(* IEC 61131-3 sources: 2026_Projet_YGO_ExcavatriceDragage/TOOLS/TEST_AUTO_CI/RESULTS/J_SUPERVISION/reports, 2 files *)

(* ---- FB_Hmi_BannerFormatter_test.st ---- *)
SETUP
VAR
    FB_Banner : FB_Hmi_BannerFormatter;
    FB_AntiFlicker : FB_AntiFlickerText;
    WinchM1Safety : ST_SafetyWinch;
    WinchM2Safety : ST_SafetyWinch;
    TranslationSafety : ST_SafetyTranslation;
    NetDiag : ST_NetworkDiagHMI;
END_VAR

// Initialisation réseau tout sain par défaut
NetDiag.InputModules.LocalDigitalIoOk := TRUE;
NetDiag.InputModules.Vh0800EndOk := TRUE;
NetDiag.InputModules.Vh0808EtpOk := TRUE;
NetDiag.InputModules.Vh0008ErOk := TRUE;
NetDiag.InputModules.Vh0008Er1Ok := TRUE;
NetDiag.BusCanOpen.Operational := TRUE;
NetDiag.Joystick.Operational := TRUE;
NetDiag.BusEthercat.Operational := TRUE;
NetDiag.EncoderM1.Operational := TRUE;
NetDiag.EncoderM2.Operational := TRUE;
NetDiag.VariateurM3.Operational := TRUE;
END_SETUP

TEST 'TC-P03-001 Dynamique Enable : neutralisation initiale, transition Ready au repos, puis coupure'
    (* Scan 0 : Enable=FALSE -> Neutralisation *)
    FB_Banner(Enable := FALSE, CurrentMode := E_Mode.DISABLE,
              EmergencyChainClosed := FALSE, PowerContactorEngaged := FALSE,
              WinchM1Safety := WinchM1Safety, WinchM2Safety := WinchM2Safety,
              Network := NetDiag);
    ASSERT_EQ(FB_Banner.Banner.GlobalContextText, '', 'Enable=FALSE -> texte vide');

    (* Scan 1 : Enable=TRUE -> Demarrage boot *)
    FB_Banner(Enable := TRUE, CurrentMode := E_Mode.MAINT_N1,
              EmergencyChainClosed := TRUE, PowerContactorEngaged := TRUE,
              WinchM1Safety := WinchM1Safety, WinchM2Safety := WinchM2Safety,
              Network := NetDiag);

    ADVANCE_TIME(5000000000); // 5s pour depasser le BootInhibit (4s)

    (* Scan 2 : Formatage actif post-boot *)
    FB_Banner(Enable := TRUE, CurrentMode := E_Mode.MAINT_N1,
              EmergencyChainClosed := TRUE, PowerContactorEngaged := TRUE,
              WinchM1Safety := WinchM1Safety, WinchM2Safety := WinchM2Safety,
              Network := NetDiag);
    ASSERT_FALSE(FB_Banner.Banner.GlobalContextText = '', 'Enable=TRUE -> non vide (nominal)');

    ADVANCE_TIME(10000000);

    (* Scan 3 : Enable=FALSE -> Re-neutralisation *)
    FB_Banner(Enable := FALSE, CurrentMode := E_Mode.DISABLE,
              EmergencyChainClosed := FALSE, PowerContactorEngaged := FALSE,
              WinchM1Safety := WinchM1Safety, WinchM2Safety := WinchM2Safety,
              Network := NetDiag);
    ASSERT_EQ(FB_Banner.Banner.GlobalContextText, '', 'Coupure -> retombe a texte vide');
END_TEST

TEST 'TC-P07-001 BannerFormatter : formatage nominal bandeau synoptique IHM'
    FB_Banner(
        Enable := TRUE,
        CurrentMode := E_Mode.MAINT_N1,
        EmergencyChainClosed := TRUE,
        PowerContactorEngaged := TRUE,
        WinchM1Safety := WinchM1Safety,
        WinchM2Safety := WinchM2Safety,
        Network := NetDiag
    );
    ADVANCE_TIME(5000000000); // 5s BootInhibit
    FB_Banner(
        Enable := TRUE,
        CurrentMode := E_Mode.MAINT_N1,
        EmergencyChainClosed := TRUE,
        PowerContactorEngaged := TRUE,
        WinchM1Safety := WinchM1Safety,
        WinchM2Safety := WinchM2Safety,
        Network := NetDiag
    );
    ASSERT_FALSE(FB_Banner.Banner.GlobalContextText = '', 'GlobalContextText non vide');
END_TEST

TEST 'TC-P07-010 AntiFlickerText : affichage instantane force'
    FB_AntiFlicker(NewText := 'TEST_INSTANT', ForceInstant := TRUE);
    ASSERT_EQ(FB_AntiFlicker.Text, 'TEST_INSTANT', 'Texte instantane');
END_TEST

TEST 'TC-P07-020 RootCause : alarme fille visible quand materiel sain'
    // Boot initial
    FB_Banner(Enable := TRUE, CurrentMode := E_Mode.MAINT_N1,
              EmergencyChainClosed := TRUE, PowerContactorEngaged := TRUE,
              WinchM1Safety := WinchM1Safety, WinchM2Safety := WinchM2Safety,
              Network := NetDiag);
    ADVANCE_TIME(5000000000); // 5s BootInhibit

    WinchM1Safety.SlackCable := TRUE; // Defaut mou de cable sur DI physique LocalDigitalIO
    FB_Banner(
        Enable := TRUE,
        CurrentMode := E_Mode.MAINT_N1,
        EmergencyChainClosed := TRUE,
        PowerContactorEngaged := TRUE,
        WinchM1Safety := WinchM1Safety,
        WinchM2Safety := WinchM2Safety,
        Network := NetDiag
    );
    ASSERT_TRUE(FB_Banner.Banner.AlarmBanner.HasAlarm, 'Alarme presente');
    ASSERT_EQ(FB_Banner.Banner.AlarmBanner.Count, 1, '1 alarme au carrousel');
    ASSERT_EQ(FB_Banner.Banner.AlarmBanner.Text, '1/1 [M1] mou de cable', 'Alarme fille correctement affichee');
    ASSERT_EQ(FB_Banner.Banner.AlarmBanner.AlarmArray[0], '[M1] mou de cable', 'Tableau AlarmArray[0] correctement rempli');
END_TEST

TEST 'TC-P07-021 RootCause : masquage alarme fille sur panne module Local_Digital_IO'
    // Boot initial
    FB_Banner(Enable := TRUE, CurrentMode := E_Mode.MAINT_N1,
              EmergencyChainClosed := TRUE, PowerContactorEngaged := TRUE,
              WinchM1Safety := WinchM1Safety, WinchM2Safety := WinchM2Safety,
              Network := NetDiag);
    ADVANCE_TIME(5000000000); // 5s BootInhibit

    WinchM1Safety.SlackCable := TRUE; // Mou de cable remonte (etat fail-safe du module HS)
    NetDiag.InputModules.LocalDigitalIoOk := FALSE; // Panne materielle coupleur/carte Local IO

    FB_Banner(
        Enable := TRUE,
        CurrentMode := E_Mode.MAINT_N1,
        EmergencyChainClosed := TRUE,
        PowerContactorEngaged := TRUE,
        WinchM1Safety := WinchM1Safety,
        WinchM2Safety := WinchM2Safety,
        Network := NetDiag
    );

    // L'alarme fille doit etre masquee, seule l'alarme parente doit apparaitre
    ASSERT_TRUE(FB_Banner.Banner.AlarmBanner.HasAlarm, 'Alarme presente');
    ASSERT_EQ(FB_Banner.Banner.AlarmBanner.Count, 1, '1 alarme (parent seul)');
    ASSERT_EQ(FB_Banner.Banner.AlarmBanner.Text, '1/1 [IO] Defaut module Local IO (DI8/DO8)', 'Alarme parente affichee');
    ASSERT_EQ(FB_Banner.Banner.AlarmBanner.AlarmArray[0], '[IO] Defaut module Local IO (DI8/DO8)', 'AlarmArray[0] porte le parent');
    ASSERT_EQ(FB_Banner.Banner.OperatorActionText, '[IO] Défaut module E/S - vérifier alimentation/coupleur', 'Consigne operateur cible la panne materielle');
END_TEST

TEST 'TC-P07-022 RootCause : masquage alarme fille sur panne module VH0800END'
    // Boot initial
    FB_Banner(Enable := TRUE, CurrentMode := E_Mode.MAINT_N1,
              EmergencyChainClosed := TRUE, PowerContactorEngaged := TRUE,
              WinchM1Safety := WinchM1Safety, WinchM2Safety := WinchM2Safety,
              Network := NetDiag);
    ADVANCE_TIME(5000000000); // 5s BootInhibit

    WinchM1Safety.ErrorPhaseRotation := TRUE;
    WinchM1Safety.ErrorBrakeThermal := TRUE;
    NetDiag.InputModules.Vh0800EndOk := FALSE; // Panne module VH0800

    FB_Banner(
        Enable := TRUE,
        CurrentMode := E_Mode.MAINT_N1,
        EmergencyChainClosed := TRUE,
        PowerContactorEngaged := TRUE,
        WinchM1Safety := WinchM1Safety,
        WinchM2Safety := WinchM2Safety,
        Network := NetDiag
    );

    ASSERT_TRUE(FB_Banner.Banner.AlarmBanner.HasAlarm, 'Alarme presente');
    ASSERT_EQ(FB_Banner.Banner.AlarmBanner.Count, 1, '1 alarme (parent seul)');
    ASSERT_EQ(FB_Banner.Banner.AlarmBanner.Text, '1/1 [IO] Defaut module VH0800END (DI8)', 'Alarme parente VH0800');
END_TEST

TEST 'TC-P07-023 RootCause : masquage alarme fille sur perte codeur ECAT'
    // Boot initial
    FB_Banner(Enable := TRUE, CurrentMode := E_Mode.MAINT_N1,
              EmergencyChainClosed := TRUE, PowerContactorEngaged := TRUE,
              WinchM1Safety := WinchM1Safety, WinchM2Safety := WinchM2Safety,
              Network := NetDiag);
    ADVANCE_TIME(5000000000); // 5s BootInhibit

    WinchM1Safety.ErrorEncoder := TRUE;
    WinchM1Safety.CableLimitDescent := TRUE;
    NetDiag.EncoderM1.Operational := FALSE; // Perte com EtherCAT codeur M1

    FB_Banner(
        Enable := TRUE,
        CurrentMode := E_Mode.MAINT_N1,
        EmergencyChainClosed := TRUE,
        PowerContactorEngaged := TRUE,
        WinchM1Safety := WinchM1Safety,
        WinchM2Safety := WinchM2Safety,
        Network := NetDiag
    );

    ASSERT_TRUE(FB_Banner.Banner.AlarmBanner.HasAlarm, 'Alarme presente');
    ASSERT_EQ(FB_Banner.Banner.AlarmBanner.Count, 1, '1 alarme (parent seul)');
    ASSERT_EQ(FB_Banner.Banner.AlarmBanner.Text, '1/1 [M1] Codeur absolu COD1 non detecte (ECAT)', 'Alarme parente codeur M1');
    ASSERT_EQ(FB_Banner.Banner.OperatorActionText, '[ECAT] Codeurs non détectés - vérifier liaison', 'Action operateur codeurs');
END_TEST

TEST 'TC-P07-024 Priorite absolue AU sur defaut module E/S'
    // Boot initial
    FB_Banner(Enable := TRUE, CurrentMode := E_Mode.MAINT_N1,
              EmergencyChainClosed := TRUE, PowerContactorEngaged := TRUE,
              WinchM1Safety := WinchM1Safety, WinchM2Safety := WinchM2Safety,
              Network := NetDiag);
    ADVANCE_TIME(5000000000); // 5s BootInhibit

    NetDiag.InputModules.LocalDigitalIoOk := FALSE;

    FB_Banner(
        Enable := TRUE,
        CurrentMode := E_Mode.MAINT_N1,
        EmergencyChainClosed := FALSE, // AU ouvert
        PowerContactorEngaged := TRUE,
        WinchM1Safety := WinchM1Safety,
        WinchM2Safety := WinchM2Safety,
        Network := NetDiag
    );

    // L'AU reste prioritaire dans la consigne operateur
    ASSERT_EQ(FB_Banner.Banner.OperatorActionText, '[PUPITRE] Boucle urgence ouverte - réarmer', 'AU domine le defaut E/S');
END_TEST

(* =======================================================================
   TC-P07-002..009 — Interface IHM (AF_Partie-07_Interface_IHM_v2.2.md §table).
   TC-P07-006/008/009 sont testables boîte noire sur FB_Hmi_BannerFormatter.
   TC-P07-002/003/004/005/007 sont des invariants structurels documentés
   (vérifiés par G200_check_linkage.py / encapsulation_check.py), pas des
   comportements runtime.
   ======================================================================= *)

TEST 'TC-P07-009 Aucun defaut actif -> bandeau d alarme vide'
    // Boot initial (reseau sain)
    FB_Banner(Enable := TRUE, CurrentMode := E_Mode.MAINT_N1,
              EmergencyChainClosed := TRUE, PowerContactorEngaged := TRUE,
              WinchM1Safety := WinchM1Safety, WinchM2Safety := WinchM2Safety,
              Network := NetDiag);
    ADVANCE_TIME(5000000000); // 5s BootInhibit

    FB_Banner(Enable := TRUE, CurrentMode := E_Mode.MAINT_N1,
              EmergencyChainClosed := TRUE, PowerContactorEngaged := TRUE,
              WinchM1Safety := WinchM1Safety, WinchM2Safety := WinchM2Safety,
              Network := NetDiag);
    ASSERT_FALSE(FB_Banner.Banner.AlarmBanner.HasAlarm, 'aucun defaut -> HasAlarm=FALSE');
    ASSERT_EQ(FB_Banner.Banner.AlarmBanner.Text, '', 'aucun defaut -> Text vide');
    ASSERT_EQ(FB_Banner.Banner.AlarmBanner.Index, 0, 'aucun defaut -> Index=0');
    ASSERT_EQ(FB_Banner.Banner.AlarmBanner.Count, 0, 'aucun defaut -> Count=0');
END_TEST

TEST 'TC-P07-008 Carrousel d alarmes : un message a la fois, index n/N coherent'
    // Boot initial (reseau sain)
    FB_Banner(Enable := TRUE, CurrentMode := E_Mode.MAINT_N1,
              EmergencyChainClosed := TRUE, PowerContactorEngaged := TRUE,
              WinchM1Safety := WinchM1Safety, WinchM2Safety := WinchM2Safety,
              Network := NetDiag);
    ADVANCE_TIME(5000000000); // 5s BootInhibit

    // 2 alarmes actives : mou de cable M1 et M2
    WinchM1Safety.SlackCable := TRUE;
    WinchM2Safety.SlackCable := TRUE;
    FB_Banner(Enable := TRUE, CurrentMode := E_Mode.MAINT_N1,
              EmergencyChainClosed := TRUE, PowerContactorEngaged := TRUE,
              WinchM1Safety := WinchM1Safety, WinchM2Safety := WinchM2Safety,
              Network := NetDiag, AlarmHoldTime := T#1s);
    ASSERT_TRUE(FB_Banner.Banner.AlarmBanner.HasAlarm, '2 defauts -> HasAlarm=TRUE');
    ASSERT_EQ(FB_Banner.Banner.AlarmBanner.Count, 2, '2 defauts -> Count=2');
    ASSERT_EQ(FB_Banner.Banner.AlarmBanner.Index, 1, 'premier message -> Index=1');
    ASSERT_EQ(FB_Banner.Banner.AlarmBanner.Text, '1/2 [M1] mou de cable', 'premier message affiche');

    // Apres AlarmHoldTime (1s) : rotation vers le message 2
    ADVANCE_TIME(1000000000);
    FB_Banner(Enable := TRUE, CurrentMode := E_Mode.MAINT_N1,
              EmergencyChainClosed := TRUE, PowerContactorEngaged := TRUE,
              WinchM1Safety := WinchM1Safety, WinchM2Safety := WinchM2Safety,
              Network := NetDiag, AlarmHoldTime := T#1s);
    ASSERT_EQ(FB_Banner.Banner.AlarmBanner.Index, 2, 'rotation -> Index=2');
    ASSERT_EQ(FB_Banner.Banner.AlarmBanner.Text, '2/2 [M2] mou de cable', 'deuxieme message affiche');

    // Apres un nouveau AlarmHoldTime : le TON a ete reset au scan precedent (rotation
    // cyclique sur 2 scans : un scan pour re-accumuler le temps, un scan pour basculer).
    ADVANCE_TIME(1000000000);
    FB_Banner(Enable := TRUE, CurrentMode := E_Mode.MAINT_N1,
              EmergencyChainClosed := TRUE, PowerContactorEngaged := TRUE,
              WinchM1Safety := WinchM1Safety, WinchM2Safety := WinchM2Safety,
              Network := NetDiag, AlarmHoldTime := T#1s);
    ASSERT_EQ(FB_Banner.Banner.AlarmBanner.Index, 2, 'scan intermediaire : TON re-accumule, pas encore de bascule');

    // Apres un second AlarmHoldTime : bascule cyclique vers le message 1
    ADVANCE_TIME(1000000000);
    FB_Banner(Enable := TRUE, CurrentMode := E_Mode.MAINT_N1,
              EmergencyChainClosed := TRUE, PowerContactorEngaged := TRUE,
              WinchM1Safety := WinchM1Safety, WinchM2Safety := WinchM2Safety,
              Network := NetDiag, AlarmHoldTime := T#1s);
    ASSERT_EQ(FB_Banner.Banner.AlarmBanner.Index, 1, 'rotation cyclique -> retour Index=1');
    ASSERT_EQ(FB_Banner.Banner.AlarmBanner.Text, '1/2 [M1] mou de cable', 'retour au premier message');
END_TEST

TEST 'TC-P07-006 Separation messages action/etat vs alarmes : alarme dans le carrousel, contexte dans le bandeau info'
    // Boot initial (reseau sain)
    FB_Banner(Enable := TRUE, CurrentMode := E_Mode.MAINT_N1,
              EmergencyChainClosed := TRUE, PowerContactorEngaged := TRUE,
              WinchM1Safety := WinchM1Safety, WinchM2Safety := WinchM2Safety,
              Network := NetDiag);
    ADVANCE_TIME(5000000000); // 5s BootInhibit

    // Une alarme active (mou de cable M1)
    WinchM1Safety.SlackCable := TRUE;
    FB_Banner(Enable := TRUE, CurrentMode := E_Mode.MAINT_N1,
              EmergencyChainClosed := TRUE, PowerContactorEngaged := TRUE,
              WinchM1Safety := WinchM1Safety, WinchM2Safety := WinchM2Safety,
              Network := NetDiag);
    // L'alarme vit dans le carrousel (AlarmBanner), pas dans le bandeau info
    ASSERT_TRUE(FB_Banner.Banner.AlarmBanner.HasAlarm, 'alarme presente dans le carrousel');
    ASSERT_EQ(FB_Banner.Banner.AlarmBanner.Text, '1/1 [M1] mou de cable', 'alarme dans le carrousel');
    // Le bandeau info (GlobalContextText) reste un contexte, pas l'alarme
    ASSERT_FALSE(FB_Banner.Banner.GlobalContextText = '', 'contexte global non vide');
    ASSERT_FALSE(FB_Banner.Banner.GlobalContextText = FB_Banner.Banner.AlarmBanner.Text,
                 'le contexte info ne porte pas le texte d alarme (2 familles distinctes)');
END_TEST

TEST 'TC-P07-002 Structures Cmd/State/Cfg par domaine (invariant structurel)'
    (* 💻 AUTO — invariant structurel documenté. Règle AF_Partie-07 §4 : convention
       Cmd/State/Cfg/Bypass/Test respectée dans GVL_IHM. FB_Hmi_BannerFormatter
       consomme des structures publiques (ST_SafetyWinch, ST_NetworkDiagHMI, E_Mode)
       et publie ST_HmiBanner. Vérifié par G200_check_linkage.py. *)
    FB_Banner(Enable := TRUE, CurrentMode := E_Mode.MAINT_N1,
              EmergencyChainClosed := TRUE, PowerContactorEngaged := TRUE,
              WinchM1Safety := WinchM1Safety, WinchM2Safety := WinchM2Safety,
              Network := NetDiag);
    ASSERT_FALSE(FB_Banner.Banner.GlobalContextText = '', 'formateur consomme des structures publiques par domaine');
END_TEST

TEST 'TC-P07-003 IHM limitee aux variables de GVL_IHM (invariant structurel)'
    (* 💻 AUTO — invariant structurel documenté. Règle AF_Partie-07 §2 : l'IHM ne lit
       ni n'écrit les internes des FB ; elle n'accède qu'à GVL_IHM. FB_Hmi_BannerFormatter
       publie Banner : ST_HmiBanner (mappé dans GVL_IHM.Banner). Vérifié par
       G200_check_linkage.py / encapsulation_check.py. *)
    FB_Banner(Enable := TRUE, CurrentMode := E_Mode.MAINT_N1,
              EmergencyChainClosed := TRUE, PowerContactorEngaged := TRUE,
              WinchM1Safety := WinchM1Safety, WinchM2Safety := WinchM2Safety,
              Network := NetDiag);
    ASSERT_FALSE(FB_Banner.Banner.GlobalContextText = '', 'sortie publique ST_HmiBanner (frontiere GVL_IHM)');
END_TEST

TEST 'TC-P07-004 Producteur unique par champ State (invariant structurel)'
    (* 💻 AUTO — invariant structurel documenté. Règle AF_Partie-07 §2 : chaque champ
       State a un seul écrivain PLC. FB_Hmi_BannerFormatter est le producteur unique
       de Banner (ST_HmiBanner) ; il ne réécrit pas les State des autres domaines.
       Vérifié par G200_check_linkage.py. *)
    FB_Banner(Enable := TRUE, CurrentMode := E_Mode.MAINT_N1,
              EmergencyChainClosed := TRUE, PowerContactorEngaged := TRUE,
              WinchM1Safety := WinchM1Safety, WinchM2Safety := WinchM2Safety,
              Network := NetDiag);
    ASSERT_FALSE(FB_Banner.Banner.GlobalContextText = '', 'producteur unique du bandeau (Banner)');
END_TEST

TEST 'TC-P07-005 Page Troubleshooting en lecture seule (invariant structurel)'
    (* 💻 AUTO — invariant structurel documenté. Règle AF_Partie-07 §7 : le troubleshooting
       est une observation lecture seule, aucune écriture de commande/config/bypass.
       Implémenté par FB_TroubleshootingView + GVL_Troubleshooting (AF_Partie-14).
       FB_Hmi_BannerFormatter ne produit aucune commande. Vérifié par
       G200_check_linkage.py / encapsulation_check.py. *)
    FB_Banner(Enable := TRUE, CurrentMode := E_Mode.MAINT_N1,
              EmergencyChainClosed := TRUE, PowerContactorEngaged := TRUE,
              WinchM1Safety := WinchM1Safety, WinchM2Safety := WinchM2Safety,
              Network := NetDiag);
    ASSERT_FALSE(FB_Banner.Banner.GlobalContextText = '', 'formateur lecture seule, aucune commande produite');
END_TEST

TEST 'TC-P07-007 Warning auto-effacable vs Fault sur Reset (invariant structurel)'
    (* ⚡ SITE+AUTO — invariant structurel documenté. Règle AF_Partie-07 §5.3 : un warning
       s'efface seul, un Fault exige Ack (pattern Cause/Ack, CODE_QUALITY_STANDARDS §9).
       Dans le bandeau, l'anti-clignotement (FB_AntiFlickerText) maintient les warnings
       min 500ms tandis que les défauts critiques passent en direct (ForceInstant).
       Le comportement Fault/Ack est porté par le socle FB_FaultCore (test_fb_faultcore.st).
       Vérifié par encapsulation_check.py. *)
    FB_Banner(Enable := TRUE, CurrentMode := E_Mode.MAINT_N1,
              EmergencyChainClosed := TRUE, PowerContactorEngaged := TRUE,
              WinchM1Safety := WinchM1Safety, WinchM2Safety := WinchM2Safety,
              Network := NetDiag);
    ASSERT_FALSE(FB_Banner.Banner.GlobalContextText = '', 'anti-clignotement gere par FB_AntiFlickerText (invariant)');
END_TEST

(* =========================================================================
   REX 2026-08-27 — Réarmement AU échouant silencieusement à l'étape 5 (PowerCutOff).
   TC-P07-030 : preuve du correctif IHM (Bug A gating + Bug B priorité + décodage
   16#0010 en cause explicite M3 MecaA). Le comportement du FB_Safety_EmergencyManagement
   (cause 16#0010, lockout, Error=FALSE, récupération Reset) est couvert par
   TC-P01-011/012/013 dans le domaine B_AU_SECURITE.
   ========================================================================= *)

TEST 'TC-P07-030 Abandon AU 16#0010 decode en cause explicite M3 MecaA (Bug A+B)'
    // Boot initial (reseau sain)
    FB_Banner(Enable := TRUE, CurrentMode := E_Mode.MAINT_N1,
              EmergencyChainClosed := TRUE, PowerContactorEngaged := TRUE,
              WinchM1Safety := WinchM1Safety, WinchM2Safety := WinchM2Safety,
              Network := NetDiag);
    ADVANCE_TIME(5000000000); // 5s BootInhibit

    // Sequence AU en cours a l etape 5 (impulsion), contacteur pulse (PowerContactorEngaged=TRUE)
    FB_Banner(Enable := TRUE, CurrentMode := E_Mode.MAINT_N1,
              EmergencyChainClosed := TRUE, PowerContactorEngaged := TRUE,
              ArmingSeqStep := 5, LastAbortCause := 16#0000,
              WinchM1Safety := WinchM1Safety, WinchM2Safety := WinchM2Safety,
              Network := NetDiag);
    ADVANCE_TIME(10000000);

    // Abandon a l etape 5 : PowerCutOff metier (16#0010) + cause M3 MecaA active.
    // Le contacteur vient d etre pulse (PowerContactorEngaged=TRUE) : l ancien gating
    // NOT PowerContactorEngaged supprimait ce message (Bug A). Il doit maintenant s afficher,
    // et la cause 16#0010 doit etre decodee en M3 MecaA (Bug B : cause avant message generique).
    TranslationSafety.ErrorMecaA := TRUE;
    FB_Banner(Enable := TRUE, CurrentMode := E_Mode.MAINT_N1,
              EmergencyChainClosed := TRUE, PowerContactorEngaged := TRUE,
              PowerCutOffActiveAny := TRUE,
              ArmingSeqStep := 0, LastAbortCause := 16#0010,
              WinchM1Safety := WinchM1Safety, WinchM2Safety := WinchM2Safety,
              TranslationSafety := TranslationSafety,
              Network := NetDiag);
    ASSERT_EQ(FB_Banner.Banner.OperatorActionText, '[M3] MecaA (mouvement non commandé) - Reset puis réarmer',
              'cause 16#0010 decodee en M3 MecaA (Bug A+B)');
END_TEST

TEST 'TC-P07-031 AX_STAB affiche le bit defaut latche, jamais #0'
    // Etat winch explicite : aucun latch, aucun mou de cable (deterministe, tests partages).
    WinchM1Safety.LatchedId := 0; WinchM1Safety.SlackCable := FALSE;
    WinchM2Safety.LatchedId := 0; WinchM2Safety.SlackCable := FALSE;
    FB_Banner(Enable := TRUE, CurrentMode := E_Mode.SEMI_AUTO,
              EmergencyChainClosed := TRUE, PowerContactorEngaged := TRUE,
              CycleStep := E_AutoCycleStep.AX_STAB,
              CycleStepAtError := E_AutoCycleStep.AX7_SEARCH_BOTTOM,
              CycleErrorId := 16#0200,
              WinchM1Safety := WinchM1Safety, WinchM2Safety := WinchM2Safety,
              Network := NetDiag);
    ASSERT_EQ(FB_Banner.Banner.OperatorActionText,
              '[CYCLE]AX7:palier 4 non confirme>Repr/Abandon',
              'AX_STAB decode le code cause cycle latche (format concis)');
END_TEST

TEST 'TC-P07-032 AX_STAB remonte la cause RACINE winch et prime sur le SafeStop generique'
    // Cause racine = vue LATCHEE (M2 MecaE). SafeStopActive est TRUE car toute cause winch
    // Meca* est une cause SafeStop : le message de cause doit malgre tout etre affiche
    // (la coupure/SafeStop est une CONSEQUENCE, pas la cause). REX 2026-09-19.
    WinchM1Safety.LatchedId := 0; WinchM1Safety.SlackCable := FALSE;
    WinchM2Safety.LatchedId := 16#3000; WinchM2Safety.SlackCable := FALSE;
    FB_Banner(Enable := TRUE, CurrentMode := E_Mode.SEMI_AUTO,
              EmergencyChainClosed := TRUE, PowerContactorEngaged := TRUE,
              SafeStopActive := TRUE,
              CycleStep := E_AutoCycleStep.AX_STAB,
              CycleStepAtError := E_AutoCycleStep.AX7_SEARCH_BOTTOM,
              CycleErrorId := 16#0200,
              WinchM1Safety := WinchM1Safety, WinchM2Safety := WinchM2Safety,
              Network := NetDiag);
    ASSERT_EQ(FB_Banner.Banner.OperatorActionText,
              '[CYCLE]AX7:palier 4 non confirme (M2 MecaE)>Repr/Abandon',
              'cause racine winch latchee affichee et prioritaire sur le message SafeStop generique');
    ASSERT_EQ(FB_Banner.Banner.SequenceProgressText,
              'Cycle: STABILISATION (defaut a AX7)',
              'repli AX_STAB : la progression situe lorigine sans laisser croire quon y est encore');
END_TEST

TEST 'TC-P07-040 T255-D limite basse cable M1 : alarme au carrousel ET action autorisee'
    // Cause VIVE non latchee (bit6 = 16#0040, FB_Safety_Winch.st:318-325) : elle allume
    // AnyFaultActive via Safety.Error mais n'etait decodee nulle part avant T255-D.
    WinchM1Safety.LatchedId := 0; WinchM1Safety.SlackCable := FALSE;
    WinchM1Safety.CableLimitDescent := TRUE;
    WinchM1Safety.Error := TRUE;
    WinchM1Safety.ErrorId := 16#0040;
    WinchM1Safety.DescendPermit := FALSE;   // interlock : descente interdite
    WinchM1Safety.AscentPermit := TRUE;     // remontee = action autorisee
    WinchM2Safety.CableLimitDescent := FALSE;
    WinchM2Safety.AscentPermit := TRUE;

    // Boot puis scan utile : depasse l'anti-clignotement (500 ms), reseau sain
    // (operateur ARME et au neutre : le prerequis homme-mort ne doit pas primer ici)
    FB_Banner(Enable := TRUE, CurrentMode := E_Mode.MAINT_N1,
              EmergencyChainClosed := TRUE, PowerContactorEngaged := TRUE,
              DeadmanArmed := TRUE, JoystickAtNeutral := TRUE,
              WinchM1Safety := WinchM1Safety, WinchM2Safety := WinchM2Safety,
              Network := NetDiag);
    ADVANCE_TIME(5000000000);
    FB_Banner(Enable := TRUE, CurrentMode := E_Mode.MAINT_N1,
              EmergencyChainClosed := TRUE, PowerContactorEngaged := TRUE,
              DeadmanArmed := TRUE, JoystickAtNeutral := TRUE,
              WinchM1Safety := WinchM1Safety, WinchM2Safety := WinchM2Safety,
              Network := NetDiag);

    ASSERT_TRUE(FB_Banner.Banner.AlarmBanner.HasAlarm, 'limite basse cable M1 : alarme presente');
    ASSERT_EQ(FB_Banner.Banner.AlarmBanner.Count, 1, 'limite basse cable M1 : une seule alarme');
    ASSERT_EQ(FB_Banner.Banner.AlarmBanner.Text, '1/1 [M1] Limite basse cable atteinte',
              'libelle alarme citant le treuil M1 et la limite basse');
    ASSERT_EQ(FB_Banner.Banner.OperatorActionText, '[TREUIL] Limite basse cable M1 - remonter',
              'action autorisee indiquee sans commande de descente');
END_TEST

TEST 'TC-P07-041 T255-D limite basse cable M2 : alarme au carrousel ET action autorisee'
    WinchM2Safety.LatchedId := 0; WinchM2Safety.SlackCable := FALSE;
    WinchM2Safety.CableLimitDescent := TRUE;
    WinchM2Safety.Error := TRUE;
    WinchM2Safety.ErrorId := 16#0040;
    WinchM2Safety.DescendPermit := FALSE;
    WinchM2Safety.AscentPermit := TRUE;
    WinchM1Safety.CableLimitDescent := FALSE;
    WinchM1Safety.AscentPermit := TRUE;

    FB_Banner(Enable := TRUE, CurrentMode := E_Mode.MAINT_N1,
              EmergencyChainClosed := TRUE, PowerContactorEngaged := TRUE,
              DeadmanArmed := TRUE, JoystickAtNeutral := TRUE,
              WinchM1Safety := WinchM1Safety, WinchM2Safety := WinchM2Safety,
              Network := NetDiag);
    ADVANCE_TIME(5000000000);
    FB_Banner(Enable := TRUE, CurrentMode := E_Mode.MAINT_N1,
              EmergencyChainClosed := TRUE, PowerContactorEngaged := TRUE,
              DeadmanArmed := TRUE, JoystickAtNeutral := TRUE,
              WinchM1Safety := WinchM1Safety, WinchM2Safety := WinchM2Safety,
              Network := NetDiag);

    ASSERT_TRUE(FB_Banner.Banner.AlarmBanner.HasAlarm, 'limite basse cable M2 : alarme presente');
    ASSERT_EQ(FB_Banner.Banner.AlarmBanner.Text, '1/1 [M2] Limite basse cable atteinte',
              'libelle alarme citant le treuil M2 et la limite basse');
    ASSERT_EQ(FB_Banner.Banner.OperatorActionText, '[TREUIL] Limite basse cable M2 - remonter',
              'action autorisee indiquee pour M2');
END_TEST

TEST 'TC-P07-042 T255-D ancre : descente commandee conserve le libelle historique'
    // Non-regression de la branche historique : sous DirectionBlocked ET descente
    // commandee, le message reste « Descente interdite - Limite basse cable » et la
    // nouvelle branche d'action ne le remplace pas.
    WinchM1Safety.CableLimitDescent := TRUE;
    WinchM1Safety.Error := TRUE;
    WinchM1Safety.ErrorId := 16#0040;
    WinchM1Safety.DescendPermit := FALSE;
    WinchM1Safety.AscentPermit := TRUE;

    FB_Banner(Enable := TRUE, CurrentMode := E_Mode.MAINT_N1,
              EmergencyChainClosed := TRUE, PowerContactorEngaged := TRUE,
              BothAxesCoupled := TRUE, WinchBothMotionDirection := -1,
              DeadmanArmed := TRUE, JoystickAtNeutral := FALSE,
              WinchM1Safety := WinchM1Safety, WinchM2Safety := WinchM2Safety,
              Network := NetDiag);
    ADVANCE_TIME(5000000000);
    FB_Banner(Enable := TRUE, CurrentMode := E_Mode.MAINT_N1,
              EmergencyChainClosed := TRUE, PowerContactorEngaged := TRUE,
              BothAxesCoupled := TRUE, WinchBothMotionDirection := -1,
              DeadmanArmed := TRUE, JoystickAtNeutral := FALSE,
              WinchM1Safety := WinchM1Safety, WinchM2Safety := WinchM2Safety,
              Network := NetDiag);

    ASSERT_EQ(FB_Banner.Banner.OperatorActionText, '[TREUIL] Descente interdite - Limite basse cable',
              'descente commandee : libelle historique inchange');
END_TEST

TEST 'TC-P07-043 T255-D ancre : champ CableLimitDescent seul NE DOIT PAS produire d alarme'
    // Le champ publie par FB_WinchStateProjection est une comparaison BRUTE de position,
    // SANS bypass ni mode referencement (FB_WinchStateProjection.st:217-218/230) : sous
    // BypassCableLimitSwitch (MAINT_N2) il reste TRUE alors que la cause safety est LEVEE
    // (ErrorId bit6 = 0) et que DescendPermit est rendu (FB_Safety_Winch.st:563-565).
    // Le carrousel doit donc lire ErrorId, jamais ce champ (revue read-only 2026-09-20).
    WinchM1Safety.LatchedId := 0; WinchM1Safety.SlackCable := FALSE;
    WinchM1Safety.CableLimitDescent := TRUE;   // etat brut de projection (bypass actif)
    WinchM1Safety.Error := FALSE;              // aucun defaut safety
    WinchM1Safety.ErrorId := 16#0000;          // bit6 leve
    WinchM1Safety.DescendPermit := TRUE;       // descente autorisee
    WinchM1Safety.AscentPermit := TRUE;
    WinchM2Safety.CableLimitDescent := FALSE;

    FB_Banner(Enable := TRUE, CurrentMode := E_Mode.MAINT_N2,
              EmergencyChainClosed := TRUE, PowerContactorEngaged := TRUE,
              DeadmanArmed := TRUE, JoystickAtNeutral := TRUE,
              WinchM1Safety := WinchM1Safety, WinchM2Safety := WinchM2Safety,
              Network := NetDiag);
    ADVANCE_TIME(5000000000);
    FB_Banner(Enable := TRUE, CurrentMode := E_Mode.MAINT_N2,
              EmergencyChainClosed := TRUE, PowerContactorEngaged := TRUE,
              DeadmanArmed := TRUE, JoystickAtNeutral := TRUE,
              WinchM1Safety := WinchM1Safety, WinchM2Safety := WinchM2Safety,
              Network := NetDiag);

    ASSERT_FALSE(FB_Banner.Banner.AlarmBanner.HasAlarm,
                 'champ de projection seul : aucune alarme ne doit apparaitre (faux positif bypass)');
    ASSERT_EQ(FB_Banner.Banner.OperatorActionText, '[JOYSTICK] Armé - actionner axe',
              'aucune consigne de remontee alors que la descente est autorisee');
END_TEST

TEST 'TC-P07-044 T255-D ancre : hors mode de marche, le prerequis de mode prime sur la remontee'
    WinchM1Safety.LatchedId := 0; WinchM1Safety.SlackCable := FALSE;
    WinchM1Safety.CableLimitDescent := TRUE;
    WinchM1Safety.Error := TRUE;
    WinchM1Safety.ErrorId := 16#0040;          // cause 6 REELLEMENT active
    WinchM1Safety.DescendPermit := FALSE;
    WinchM1Safety.AscentPermit := TRUE;

    FB_Banner(Enable := TRUE, CurrentMode := E_Mode.DISABLE,
              EmergencyChainClosed := TRUE, PowerContactorEngaged := TRUE,
              DeadmanArmed := TRUE, JoystickAtNeutral := TRUE,
              WinchM1Safety := WinchM1Safety, WinchM2Safety := WinchM2Safety,
              Network := NetDiag);
    ADVANCE_TIME(5000000000);
    FB_Banner(Enable := TRUE, CurrentMode := E_Mode.DISABLE,
              EmergencyChainClosed := TRUE, PowerContactorEngaged := TRUE,
              DeadmanArmed := TRUE, JoystickAtNeutral := TRUE,
              WinchM1Safety := WinchM1Safety, WinchM2Safety := WinchM2Safety,
              Network := NetDiag);

    ASSERT_TRUE(FB_Banner.Banner.AlarmBanner.HasAlarm, 'la cause reste visible au carrousel en DISABLE');
    ASSERT_EQ(FB_Banner.Banner.OperatorActionText, '[IHM] Sélectionner un mode',
              'hors mode de marche : consigne de mode, jamais une action inexécutable');
END_TEST

(* =========================================================================
   T359 / T278 — MASQUAGE BORNE DES ALARMES RESEAU PARASITES (option O1)
   =========================================================================
   BESOIN CLIENT (mail GCAM, T278) : a chaque ouverture d'AU, demarrage CPU et
   rearmement puissance, les esclaves publient des pertes de liaison de quelques
   scans. Aujourd'hui le bandeau les affiche : le TOF anti-bagotement
   (FB_Hmi_BannerFormatter.st:197-207, PT := T#1.5s) MAINTIENT l'alarme 1,5 s,
   d'ou une cascade de faux positifs que l'operateur doit acquitter.

   CIBLE : masquer les defauts RESEAU/ES uniquement pendant une fenetre transitoire
   ou leur absence est ATTENDUE (AU ouverte, rearmement puissance, boot), et
   l'afficher normalement hors de cette fenetre. Un defaut persistant reste donc
   affiche des la fin de la fenetre : le masquage est BORNE, jamais silencieux.

   TC-T359-004 est la PREUVE AVANT CORRECTIF : elle est ROUGE sur l'etat actuel.
   TC-T359-005 verrouille la BORNE (le masque ne peut pas cacher un defaut durable).
   TC-T359-006 verrouille la non-regression safety (la cause AU reste prioritaire).
   ========================================================================= *)

TEST 'TC-T359-004 Fenetre de rearmement : les pertes de liaison transitoires ne sont PAS affichees'
    (* Scan 0 : AU fermee, contacteur AU REPOS -> garde de demarrage lancee *)
    FB_Banner(Enable := TRUE, CurrentMode := E_Mode.MAINT_N1,
              EmergencyChainClosed := TRUE, PowerContactorEngaged := FALSE,
              WinchM1Safety := WinchM1Safety, WinchM2Safety := WinchM2Safety,
              Network := NetDiag);
    ASSERT_FALSE(FB_Banner.Banner.AlarmBanner.HasAlarm, 'Depart : aucune alarme');

    (* Sortie de la garde de demarrage : 4 s ecoulees, contacteur toujours au repos *)
    ADVANCE_TIME(5000000000);
    FB_Banner(Enable := TRUE, CurrentMode := E_Mode.MAINT_N1,
              EmergencyChainClosed := TRUE, PowerContactorEngaged := FALSE,
              WinchM1Safety := WinchM1Safety, WinchM2Safety := WinchM2Safety,
              Network := NetDiag);
    ASSERT_FALSE(FB_Banner.Banner.AlarmBanner.HasAlarm, 'Garde de demarrage ecoulee, reseau sain');

    (* REARMEMENT PUISSANCE : front du contacteur -> fenetre transitoire bornee ouverte *)
    FB_Banner(Enable := TRUE, CurrentMode := E_Mode.MAINT_N1,
              EmergencyChainClosed := TRUE, PowerContactorEngaged := TRUE,
              WinchM1Safety := WinchM1Safety, WinchM2Safety := WinchM2Safety,
              Network := NetDiag);

    (* Les esclaves ne sont PAS encore operationnels : c'est le transitoire reel machine *)
    NetDiag.BusEthercat.Operational := FALSE;
    NetDiag.EncoderM1.Operational := FALSE;
    NetDiag.EncoderM2.Operational := FALSE;

    ADVANCE_TIME(100000000); // 100 ms : largement au-dela d'un scan, tres en deca de 1,5 s
    FB_Banner(Enable := TRUE, CurrentMode := E_Mode.MAINT_N1,
              EmergencyChainClosed := TRUE, PowerContactorEngaged := TRUE,
              WinchM1Safety := WinchM1Safety, WinchM2Safety := WinchM2Safety,
              Network := NetDiag);

    (* CIBLE T278 : aucune alarme parasite pendant la fenetre de rearmement *)
    ASSERT_FALSE(FB_Banner.Banner.AlarmBanner.HasAlarm,
                 'Fenetre de rearmement : aucune alarme reseau parasite (cible T278)');
END_TEST

TEST 'TC-T359-005 Borne du masquage : un defaut reseau durable EST affiche des la fin de la fenetre'
    (* Meme sequence que TC-T359-004 : rearmement puis perte de liaison *)
    FB_Banner(Enable := TRUE, CurrentMode := E_Mode.MAINT_N1,
              EmergencyChainClosed := TRUE, PowerContactorEngaged := FALSE,
              WinchM1Safety := WinchM1Safety, WinchM2Safety := WinchM2Safety,
              Network := NetDiag);
    ADVANCE_TIME(5000000000);
    FB_Banner(Enable := TRUE, CurrentMode := E_Mode.MAINT_N1,
              EmergencyChainClosed := TRUE, PowerContactorEngaged := TRUE,
              WinchM1Safety := WinchM1Safety, WinchM2Safety := WinchM2Safety,
              Network := NetDiag);

    NetDiag.BusEthercat.Operational := FALSE;
    ADVANCE_TIME(100000000);
    FB_Banner(Enable := TRUE, CurrentMode := E_Mode.MAINT_N1,
              EmergencyChainClosed := TRUE, PowerContactorEngaged := TRUE,
              WinchM1Safety := WinchM1Safety, WinchM2Safety := WinchM2Safety,
              Network := NetDiag);

    (* La fenetre se referme : le defaut TOUJOURS present doit reapparaitre.
       Sans cette borne, le masquage cacherait une panne reelle de facon permanente. *)
    ADVANCE_TIME(10000000000); // 10 s : bien au-dela de toute fenetre transitoire
    FB_Banner(Enable := TRUE, CurrentMode := E_Mode.MAINT_N1,
              EmergencyChainClosed := TRUE, PowerContactorEngaged := TRUE,
              WinchM1Safety := WinchM1Safety, WinchM2Safety := WinchM2Safety,
              Network := NetDiag);

    ASSERT_TRUE(FB_Banner.Banner.AlarmBanner.HasAlarm,
                'Apres la fenetre : un defaut reseau PERSISTANT est affiche');
    ASSERT_EQ(FB_Banner.Banner.AlarmBanner.Text, '1/1 [ECAT] Defaut bus EtherCAT',
              'Le defaut durable affiche est bien celui du bus EtherCAT');
END_TEST

TEST 'TC-T359-006 Non-regression safety : la cause AU reste prioritaire, jamais masquee'
    (* AU ouverte + defaut de bus : le masquage reseau ne doit JAMAIS toucher la cause safety *)
    FB_Banner(Enable := TRUE, CurrentMode := E_Mode.MAINT_N1,
              EmergencyChainClosed := TRUE, PowerContactorEngaged := TRUE,
              WinchM1Safety := WinchM1Safety, WinchM2Safety := WinchM2Safety,
              Network := NetDiag);
    ADVANCE_TIME(5000000000);

    NetDiag.BusEthercat.Operational := FALSE;
    FB_Banner(Enable := TRUE, CurrentMode := E_Mode.MAINT_N1,
              EmergencyChainClosed := FALSE, // AU ouverte : cause safety
              PowerContactorEngaged := TRUE,
              WinchM1Safety := WinchM1Safety, WinchM2Safety := WinchM2Safety,
              Network := NetDiag);

    ASSERT_EQ(FB_Banner.Banner.OperatorActionText, '[PUPITRE] Boucle urgence ouverte - réarmer',
              'La consigne operateur reste la cause AU malgre le defaut de bus');
END_TEST

(* ═══════════════════════════════════════════════════════════════════════════════
   T368 - TEMPS ECOULE DU CYCLE ACCOLE AU BANDEAU MODE (format MMminSSs)
   Contrat : DOC/WFLOW/CONTRACTS/TASK_CONTRACT_T368_TEMPS_ECOULE_BANDEAU_AX13.yaml (AC1, AC2).
   Le suffixe n apparait QUE pendant un cycle reellement en cours (CycleAutoBusy = Lifecycle.Busy
   du sequenceur, cable PRG_07_Supervision.st:758) : hors cycle, aucune duree figee n est
   affichee. Les deux valeurs arrivent par VAR_INPUT : le formateur ne lit aucun global.
   ═══════════════════════════════════════════════════════════════════════════════ *)

TEST 'T368-001 : bandeau mode porteur du temps ecoule, uniquement pendant un cycle en cours'
    FB_Banner(Enable := TRUE, SimulationModeActive := TRUE, CurrentMode := E_Mode.SEMI_AUTO,
              CycleAutoBusy := TRUE, CycleElapsed_Min := 0, CycleElapsed_S := 0,
              EmergencyChainClosed := TRUE, PowerContactorEngaged := TRUE,
              WinchM1Safety := WinchM1Safety, WinchM2Safety := WinchM2Safety,
              Network := NetDiag);
    ADVANCE_TIME(5000000000);

    (* Scan 1 : cycle en cours, chrono a zero -> le suffixe zero-padde est present. *)
    FB_Banner(Enable := TRUE, SimulationModeActive := TRUE, CurrentMode := E_Mode.SEMI_AUTO,
              CycleAutoBusy := TRUE, CycleElapsed_Min := 0, CycleElapsed_S := 0,
              EmergencyChainClosed := TRUE, PowerContactorEngaged := TRUE,
              WinchM1Safety := WinchM1Safety, WinchM2Safety := WinchM2Safety,
              Network := NetDiag);
    ASSERT_EQ(FB_Banner.Banner.GlobalContextText, '[SIMULATION] [SEMI-AUTO] [CYCLE AUTO] 00min00s',
              'T368 : cycle en cours -> bandeau mode suivi du chrono MMminSSs');

    (* Scan 2 : 1 min 05 s -> chaque champ garde 2 chiffres (00min05s vs 1min5s : discriminant). *)
    FB_Banner(Enable := TRUE, SimulationModeActive := TRUE, CurrentMode := E_Mode.SEMI_AUTO,
              CycleAutoBusy := TRUE, CycleElapsed_Min := 1, CycleElapsed_S := 5,
              EmergencyChainClosed := TRUE, PowerContactorEngaged := TRUE,
              WinchM1Safety := WinchM1Safety, WinchM2Safety := WinchM2Safety,
              Network := NetDiag);
    ASSERT_EQ(FB_Banner.Banner.GlobalContextText, '[SIMULATION] [SEMI-AUTO] [CYCLE AUTO] 01min05s',
              'T368 : minutes et secondes zero-paddees (01min05s), aucun champ a 1 chiffre');

    (* Scan 3 : cycle termine (Busy retombe) -> bandeau mode STRICTEMENT nu, aucune duree figee. *)
    FB_Banner(Enable := TRUE, SimulationModeActive := TRUE, CurrentMode := E_Mode.SEMI_AUTO,
              CycleAutoBusy := FALSE, CycleElapsed_Min := 1, CycleElapsed_S := 5,
              EmergencyChainClosed := TRUE, PowerContactorEngaged := TRUE,
              WinchM1Safety := WinchM1Safety, WinchM2Safety := WinchM2Safety,
              Network := NetDiag);
    ASSERT_EQ(FB_Banner.Banner.GlobalContextText, '[SIMULATION] [SEMI-AUTO] [CYCLE AUTO]',
              'T368 : hors cycle -> aucune duree affichee, meme si les entrees portent encore 1 min 05 s');
END_TEST

(* ---- FB_TroubleshootingView_test.st ---- *)
(* =======================================================================
   🧪 test_fb_troubleshootingview.st — FB_TroubleshootingView (TC-P14-TSV-01..05)
   ───────────────────────────────────────────────────────────────
   Lot : écriture de tests CI — domaine AF-14 (troubleshooting).
   Fiche : DOC/AF/AF_Partie-14_Fonction_Troubleshooting/FB_TroubleshootingView_v1.2.md §8.
   Conventions : 1 appel FB() = 1 scan. Le FB est lecture-pure : il recopie des faits
   déjà publiés vers GVL_Troubleshooting (aucune commande). Les scénarios assertent
   sur les valeurs d'init sûres de GVL_Troubleshooting.* et sur l'interface (Ready).
   Les TC de pure architecture (G200, gates) portent une assertion d'invariant
   structurel documenté + commentaire « (essai d'architecture — validation partielle
   boîte noire) ».
   ======================================================================= *)

SETUP
VAR
    FB : FB_TroubleshootingView;
END_VAR
END_SETUP

TEST 'TC-P14-TSV-01 Interface : seule sortie Ready, aucune commande (essai d architecture - validation partielle boite noire)'
    (* Enable=FALSE -> Ready=FALSE (neutralisation) *)
    FB(Enable := FALSE);
    ASSERT_FALSE(FB.Ready, 'Enable=FALSE -> Ready=FALSE');

    (* Enable=TRUE -> Ready=TRUE *)
    FB(Enable := TRUE);
    ASSERT_TRUE(FB.Ready, 'Enable=TRUE -> Ready=TRUE');

    (* (essai d architecture - validation partielle boite noire) : l interface VAR_OUTPUT de
       FB_TroubleshootingView = Ready uniquement (fiche §3) -- aucune sortie SafeStop/Enable/
       Cmd/Bypass/Config. Toute publication passe par GVL_Troubleshooting (lecture seule). *)
END_TEST

TEST 'TC-P14-TSV-02 Chaque champ GVL_Troubleshooting a un producteur documente : init sure (essai d architecture - validation partielle boite noire)'
    (* Appel nominal : tous les inputs par defaut (FALSE/0) -> le FB recopie les faits
       publies vers GVL_Troubleshooting. On verifie l initialisation sure des champs. *)
    FB(Enable := TRUE);
    ASSERT_EQ(GVL_Troubleshooting.A_ContexteMachineGlobal.Idx101_ModeActive, E_Mode.DISABLE,
              'Idx101_ModeActive = Auth.Mode (init DISABLE)');
    ASSERT_FALSE(GVL_Troubleshooting.A_ContexteMachineGlobal.Idx102_SimulationEnabled,
                 'Idx102_SimulationEnabled = FALSE (init)');
    ASSERT_FALSE(GVL_Troubleshooting.A_ContexteMachineGlobal.Idx202_BypassNetworkGlobal,
                 'Idx202_BypassNetworkGlobal = FALSE (init)');
    ASSERT_FALSE(GVL_Troubleshooting.A_ContexteMachineGlobal.Idx401_HmiHeartbeatOk,
                 'Idx401_HmiHeartbeatOk = FALSE (init)');
    ASSERT_FALSE(GVL_Troubleshooting.H_LevageSynchroniseM1M2.Idx302_SyncFaultActive,
                 'Idx302_SyncFaultActive = FALSE (init)');
END_TEST

TEST 'TC-P14-TSV-03 Champs TBD publies a leur valeur d init (aucune mesure inventee)'
    (* Fiche §6/§7 : un champ sans producteur reel reste a sa valeur d initialisation,
       jamais recalculé. On verifie les 4 champs TBD documentes. *)
    FB(Enable := TRUE);
    ASSERT_FALSE(GVL_Troubleshooting.A_ContexteMachineGlobal.Idx203_BypassSensorsGlobal,
                 'Idx203_BypassSensorsGlobal = FALSE (TBD non cable)');
    ASSERT_FALSE(GVL_Troubleshooting.I_LevageUnitaireM1.Safety_300.Idx307_SlackCablePhysical_DI,
                 'Idx307_SlackCablePhysical_DI = FALSE (TBD)');
    ASSERT_FALSE(GVL_Troubleshooting.K_BenneOuvertureFermeture.Idx501_M2_CmdRev_DQ,
                 'Idx501_M2_CmdRev_DQ = FALSE (TBD)');
    ASSERT_EQ(GVL_Troubleshooting.L_TranslationPontM3.Outputs_500.Idx502_CmdDriveFreq_Hz, 0,
             'Idx502_CmdDriveFreq_Hz = 0 (TBD)');
END_TEST

TEST 'TC-P14-TSV-04 Instance unique appelee dans PRG_07_Supervision (G200) (essai d architecture - validation partielle boite noire)'
    (* (essai d architecture - validation partielle boite noire) : la liaison G200 (instance
       unique, appelee dans PRG_07_Supervision seul) est verifiee par G200_check_linkage.py,
       pas par le harnais. Ce scenario verifie que le FB est fonctionnel en boite noire. *)
    FB(Enable := TRUE);
    ASSERT_TRUE(FB.Ready, 'FB_TroubleshootingView pret (lecture seule)');
END_TEST

TEST 'TC-P14-TSV-05 Aucune regression gates (essai d architecture - validation partielle boite noire)'
    (* (essai d architecture - validation partielle boite noire) : la non-regression des gates
       est verifiee par run_all_gates.py, pas par le harnais. Scenario logique minimal. *)
    FB(Enable := TRUE);
    ASSERT_TRUE(FB.Ready, 'FB_TroubleshootingView pret');
END_TEST

(* =======================================================================
   🛡️ T371 — FAUX VERT DU DIAGNOSTIC MOUVEMENT (Step8_OutputInterlockOk)
   ───────────────────────────────────────────────────────────────
   ⚠️ COMMENT CE FB EST ALIMENTE EN TEST : FB_TroubleshootingView est LECTURE-PURE. Il recopie des
   faits DEJA PUBLIES par d'autres (GVL_IHM / GVL_Troubleshooting) : les scenarios ci-dessous pilotent
   donc ses ENTREES (`FB.WinchM1`, `FB.WinchM2`, `FB.Translation`) avec les valeurs REELLES que la
   barriere finale produit — elles ne sont pas inventees, elles sont citees ligne a ligne ci-dessous.
   La barriere (FB_WinchOutputInterlock) n'est PAS dans la chaine de compilation de ce harnais : elle
   ne peut donc pas etre pilotee ici, et ces cas ne la pilotent pas.

   📌 LES 4 MODES DE REFUS A FAUX VERT (preuve statique, FB_WinchOutputInterlock.st) :
     F1 :357-363  RestartInhibit                       -> State FAULT,              Reason RESTART_INHIBITED
     F2 :364-373  ContactorStuckLatched                -> State FAULT,              Reason SENSE_DROP_TIMEOUT
     F3 :393-404  SafeStop OU PermitFinalBlocked       -> State READY (!),          Reason NONE (!)
     F4 :424-429  RestartRequired OU DeadTimePending   -> State WAIT_RESTART_DELAY, Reason NONE (!)
   Dans les 4 cas Fault.Error = FALSE (cause unique = ErrorId bit0, timeout frein, :516-519 -> :528-532) :
   l'ancien `Step8 := NOT FinalInterlockError` (:577/:609/:644) rendait donc TRUE = FAUX VERT.

   ⚠️ HONNETETE SUR CE QUI EST PROUVE ICI : seule la barriere est fautive sur `Step8`.
   `AllConditionsMet` etait DEJA FALSE dans les 4 modes, par `Step7_BrakeReleased` (= BrakeCmd AND
   BrakeCommandOpenConfirmed) : la barriere coupe BrakeCmd (= RelayFwd OR RelayRev) dans tous ces
   refus, donc Step7 tombe a FALSE et l'ET se propage. Ces cas n'assertent donc PAS AllConditionsMet
   (le faire serait vacue) : ils assertent le seul champ qui mentait, Step8.

   ⚠️ ETAT D'EXECUTION (2026-09-21, T371) : ces cas SONT EXECUTES (ROUGE mesure avant correctif, VERT apres).
   Les DEUX murs PREEXISTANTS a HEAD qui les rendaient non jouables ont ete leves par T371 :
     (1) 8 types manquants dans l'entree `FB_TroubleshootingView` de registry.yaml — CORRIGE (8 lignes) ;
     (2) STruCpp v0.6.2 ne supporte PAS le namespace GVL de CODESYS (`GVL_Troubleshooting.X`) :
         levee par 2 MOCKS miroirs (`TOOLS/TEST_AUTO_CI/MOCKS/MOCK_GVL_*.st`) qui declarent
         `GVL_Troubleshooting` / `GVL_IHM` comme VARIABLES globales de STRUCT miroirs.
   ⚠️ REALISME DES VALEURS PILOTEES (REX revue independante T371, verdict BLOCK du 2026-09-21) : dans un
   refus, la DEMANDE reste presente (FB_Winch demande toujours) et la barriere coupe SA SORTIE. Les cas
   ci-dessous pilotent donc `RelayFwd := TRUE` (demande, miroir de FB_Winch, projection :102-103) AVEC
   `BrakeCmd := FALSE` (SORTIE validee de la barriere, projection :108). Un cas qui mettrait
   `RelayFwd := FALSE` fabriquerait un etat IMPOSSIBLE en exploitation et validerait un temoin tautologique.
   ======================================================================= *)

TEST 'TC-P14-TSV-06 M1/F1 : barriere FAULT + RESTART_INHIBITED, Fault.Error=FALSE -> Step8 PAS vert'
    (* Valeurs publiees par la barriere au site F1 (:357-363), projetees par FB_WinchStateProjection.st:112-115 *)
    FB.WinchM1.State.FinalInterlockError  := FALSE;                                    // bit0 non pose
    FB.WinchM1.State.FinalInterlockState  := E_WinchFinalInterlockState.FAULT;          // :363
    FB.WinchM1.State.FinalInterlockReason := E_WinchFinalInterlockReason.RESTART_INHIBITED; // :362
    FB.WinchM1.State.FinalMotorRequest    := TRUE;                                      // :118 projection (vue barriere)
    FB.WinchM1.State.RelayFwd             := TRUE;                                      // DEMANDE (miroir FB_Winch, :102)
    FB.WinchM1.State.RelayRev             := FALSE;
    FB.WinchM1.State.BrakeCmd             := FALSE;                                     // SORTIE validee coupee (:108 -> :487)
    FB(Enable := TRUE);
    ASSERT_EQ(GVL_Troubleshooting.N_MotionM1.Step8_InterlockState, E_WinchFinalInterlockState.FAULT, 'Step8_InterlockState = FAULT');
    ASSERT_EQ(GVL_Troubleshooting.N_MotionM1.Step8_InterlockReason, E_WinchFinalInterlockReason.RESTART_INHIBITED, 'Step8_InterlockReason = RESTART_INHIBITED');
    ASSERT_FALSE(GVL_Troubleshooting.N_MotionM1.Step8_OutputInterlockOk,
                 'F1 RestartInhibit : la barriere refuse -> Step8 doit etre FALSE (faux vert avant T371)');
END_TEST

TEST 'TC-P14-TSV-07 M1/F2 : barriere FAULT + SENSE_DROP_TIMEOUT, Fault.Error=FALSE -> Step8 PAS vert'
    (* Site F2 (:364-373) — latch T_max §3bis, sans aucun defaut frein *)
    FB.WinchM1.State.FinalInterlockError  := FALSE;
    FB.WinchM1.State.FinalInterlockState  := E_WinchFinalInterlockState.FAULT;              // :373
    FB.WinchM1.State.FinalInterlockReason := E_WinchFinalInterlockReason.SENSE_DROP_TIMEOUT; // :372
    FB.WinchM1.State.FinalMotorRequest    := TRUE;
    FB.WinchM1.State.RelayFwd             := TRUE;    // demande toujours presente
    FB.WinchM1.State.RelayRev             := FALSE;
    FB.WinchM1.State.BrakeCmd             := FALSE;   // sortie validee coupee
    FB(Enable := TRUE);
    ASSERT_EQ(GVL_Troubleshooting.N_MotionM1.Step8_InterlockReason, E_WinchFinalInterlockReason.SENSE_DROP_TIMEOUT, 'Step8_InterlockReason = SENSE_DROP_TIMEOUT');
    ASSERT_FALSE(GVL_Troubleshooting.N_MotionM1.Step8_OutputInterlockOk,
                 'F2 ContactorStuckLatched : la barriere refuse -> Step8 doit etre FALSE');
END_TEST

TEST 'TC-P14-TSV-08 M1/F3 : SafeStop/PermitFinalBlocked (State=READY, Reason=NONE) -> Step8 PAS vert'
    (* Site F3 (:393-404) — LE PLUS TROMPEUR : State laisse a READY et Reason a NONE alors que les
       6 ordres sont coupes (:402-403). Etat REEL en exploitation : la demande est TOUJOURS la
       (RelayFwd = TRUE, miroir de FB_Winch) et c'est la SORTIE VALIDEE qui est coupee (BrakeCmd = FALSE).
       Ce cas est celui qui a fait tomber la 1re version du correctif (temoin tautologique sur
       RelayFwd/RelayRev, cf. REX revue independante) : il ne doit JAMAIS etre adouci. *)
    FB.WinchM1.State.FinalInterlockError  := FALSE;
    FB.WinchM1.State.FinalInterlockState  := E_WinchFinalInterlockState.READY;   // :404 — piege
    FB.WinchM1.State.FinalInterlockReason := E_WinchFinalInterlockReason.NONE;   // non ecrit
    FB.WinchM1.State.FinalMotorRequest    := TRUE;                              // demande vivante
    FB.WinchM1.State.RelayFwd             := TRUE;                              // DEMANDE presente
    FB.WinchM1.State.RelayRev             := FALSE;
    FB.WinchM1.State.BrakeCmd             := FALSE;                             // aucune sortie validee
    FB(Enable := TRUE);
    ASSERT_FALSE(GVL_Troubleshooting.N_MotionM1.Step8_OutputInterlockOk,
                 'F3 SafeStop/PermitFinalBlocked : sortie coupee -> Step8 doit etre FALSE malgre State=READY');
END_TEST

TEST 'TC-P14-TSV-09 M1/F4 : RestartRequired/DeadTimePending (WAIT_RESTART_DELAY) -> Step8 PAS vert'
    (* Site F4 (:424-429) — Reason reste NONE : un correctif lisant Reason SEUL raterait F3 et F4 *)
    FB.WinchM1.State.FinalInterlockError  := FALSE;
    FB.WinchM1.State.FinalInterlockState  := E_WinchFinalInterlockState.WAIT_RESTART_DELAY; // :429
    FB.WinchM1.State.FinalInterlockReason := E_WinchFinalInterlockReason.NONE;
    FB.WinchM1.State.FinalMotorRequest    := TRUE;
    FB.WinchM1.State.RelayFwd             := TRUE;    // demande presente
    FB.WinchM1.State.RelayRev             := FALSE;
    FB.WinchM1.State.BrakeCmd             := FALSE;   // sortie retenue par la tempo
    FB(Enable := TRUE);
    ASSERT_EQ(GVL_Troubleshooting.N_MotionM1.Step8_InterlockState, E_WinchFinalInterlockState.WAIT_RESTART_DELAY, 'Step8_InterlockState = WAIT_RESTART_DELAY');
    ASSERT_FALSE(GVL_Troubleshooting.N_MotionM1.Step8_OutputInterlockOk,
                 'F4 tempos anti-court-cycle : demande retenue -> Step8 doit etre FALSE');
END_TEST

TEST 'TC-P14-TSV-10 M2/F3 : meme patron sur l axe M2 (State=READY, sortie coupee) -> Step8 PAS vert'
    (* Source M2 : FB_WinchStateProjection.st:179-182 + FB_WinchOutputInterlock.st:393-404.
       Meme realisme que M1 : demande presente, sortie validee coupee. *)
    FB.WinchM2.State.FinalInterlockError  := FALSE;
    FB.WinchM2.State.FinalInterlockState  := E_WinchFinalInterlockState.READY;
    FB.WinchM2.State.FinalInterlockReason := E_WinchFinalInterlockReason.NONE;
    FB.WinchM2.State.FinalMotorRequest    := TRUE;
    FB.WinchM2.State.RelayFwd             := TRUE;    // demande presente (miroir FB_Winch :175)
    FB.WinchM2.State.RelayRev             := FALSE;
    FB.WinchM2.State.BrakeCmd             := FALSE;   // sortie validee coupee (projection :175)
    FB(Enable := TRUE);
    ASSERT_FALSE(GVL_Troubleshooting.O_MotionM2.Step8_OutputInterlockOk,
                 'M2 F3 : sortie coupee -> Step8 doit etre FALSE malgre State=READY');
END_TEST

TEST 'TC-P14-TSV-11 M3 : etat et cause de la barriere M3 publies, defaut = PAS vert'
    (* M3 : la barriere publie Fault.Error (source unique) + Reason (memoire). Son ordre VALIDE existe
       bien ailleurs (PRG_06:458 -> PRG_07:576 `GVL_IHM.IoHw.Out.M3_CommandWord`) mais n'est PAS une
       entree de ce FB : l'atteindre exigerait d'ajouter `IoHw` en VAR_INPUT + un argument dans
       PRG_07_Supervision.st (hors perimetre T371). Limite declaree, remontee a l'orchestrateur. *)
    FB.Translation.State.FinalInterlockError  := TRUE;   // timeout confirmation frein M3
    FB.Translation.State.FinalInterlockState  := E_State.ERROR;
    FB.Translation.State.FinalInterlockReason := E_TranslationFinalInterlockReason.BRAKE_COMMAND_NOT_CONFIRMED;
    FB(Enable := TRUE);
    ASSERT_EQ(GVL_Troubleshooting.P_MotionM3.Step8_InterlockState, E_WinchFinalInterlockState.FAULT, 'Step8_InterlockState M3 = FAULT (projete depuis E_State.ERROR)');
    ASSERT_EQ(GVL_Troubleshooting.P_MotionM3.Step8_InterlockReason, E_WinchFinalInterlockReason.BRAKE_COMMAND_NOT_CONFIRMED, 'Step8_InterlockReason M3 = BRAKE_COMMAND_NOT_CONFIRMED');
    ASSERT_FALSE(GVL_Troubleshooting.P_MotionM3.Step8_OutputInterlockOk,
                 'M3 en defaut -> Step8 doit etre FALSE');
END_TEST

TEST 'TC-P14-TSV-12 NON-REGRESSION : barriere nominale au repos -> Step8 reste VERT (pas de faux rouge)'
    (* Garde-fou anti-sur-correction : au repos (State READY, aucune demande, aucun defaut) la
       conclusion doit rester VERTE. Verifie aussi les 2 etats NON bloquants ou l'etage de sortie est
       bien engage : WAIT_BRAKE_COMMAND_CONFIRMATION (ordre emis) et WAIT_SENSE_DROP_CONFIRM (§3bis). *)
    FB.WinchM1.State.FinalInterlockError  := FALSE;
    FB.WinchM1.State.FinalInterlockReason := E_WinchFinalInterlockReason.NONE;
    FB.WinchM1.State.FinalInterlockState  := E_WinchFinalInterlockState.READY;
    FB.WinchM1.State.FinalMotorRequest    := FALSE;   // aucune demande
    FB.WinchM1.State.RelayFwd             := FALSE;
    FB.WinchM1.State.RelayRev             := FALSE;
    FB(Enable := TRUE);
    ASSERT_TRUE(GVL_Troubleshooting.N_MotionM1.Step8_OutputInterlockOk, 'Repos nominal -> Step8 = TRUE');

    FB.WinchM1.State.FinalInterlockState := E_WinchFinalInterlockState.WAIT_BRAKE_COMMAND_CONFIRMATION;
    FB.WinchM1.State.FinalMotorRequest   := TRUE;
    FB.WinchM1.State.RelayFwd            := TRUE;     // ordre de sens emis : etage de sortie engage
    FB.WinchM1.State.BrakeCmd            := TRUE;     // SORTIE validee presente -> pas un refus
    FB(Enable := TRUE);
    ASSERT_TRUE(GVL_Troubleshooting.N_MotionM1.Step8_OutputInterlockOk,
                'Attente confirmation frein (ordre emis) -> PAS un refus, Step8 = TRUE');

    FB.WinchM1.State.FinalInterlockState := E_WinchFinalInterlockState.WAIT_SENSE_DROP_CONFIRM;
    FB.WinchM1.State.FinalMotorRequest   := FALSE;    // §3bis : palier retombe, sens tenu
    FB.WinchM1.State.RelayFwd            := TRUE;
    FB(Enable := TRUE);
    ASSERT_TRUE(GVL_Troubleshooting.N_MotionM1.Step8_OutputInterlockOk,
                'Maintien §3bis du sens -> PAS un refus, Step8 = TRUE');
END_TEST

TEST 'TC-P14-TSV-13 M2/F1 : barriere FAULT + RESTART_INHIBITED (demande vivante) -> Step8 PAS vert'
    (* Complement de couverture exige par la revue independante : F1 n'etait teste que sur M1. *)
    FB.WinchM2.State.FinalInterlockError  := FALSE;
    FB.WinchM2.State.FinalInterlockState  := E_WinchFinalInterlockState.FAULT;              // :363
    FB.WinchM2.State.FinalInterlockReason := E_WinchFinalInterlockReason.RESTART_INHIBITED; // :362
    FB.WinchM2.State.FinalMotorRequest    := TRUE;
    FB.WinchM2.State.RelayFwd             := TRUE;    // demande presente
    FB.WinchM2.State.RelayRev             := FALSE;
    FB.WinchM2.State.BrakeCmd             := FALSE;   // sortie validee coupee
    FB(Enable := TRUE);
    ASSERT_FALSE(GVL_Troubleshooting.O_MotionM2.Step8_OutputInterlockOk,
                 'M2 F1 RestartInhibit : la barriere refuse -> Step8 doit etre FALSE');
END_TEST

TEST 'TC-P14-TSV-14 M2/F4 : tempos (WAIT_RESTART_DELAY), demande retenue -> Step8 PAS vert'
    (* Complement de couverture exige par la revue independante : F4 n'etait teste que sur M1. *)
    FB.WinchM2.State.FinalInterlockError  := FALSE;
    FB.WinchM2.State.FinalInterlockState  := E_WinchFinalInterlockState.WAIT_RESTART_DELAY; // :429
    FB.WinchM2.State.FinalInterlockReason := E_WinchFinalInterlockReason.NONE;
    FB.WinchM2.State.FinalMotorRequest    := TRUE;
    FB.WinchM2.State.RelayFwd             := TRUE;
    FB.WinchM2.State.RelayRev             := FALSE;
    FB.WinchM2.State.BrakeCmd             := FALSE;
    FB(Enable := TRUE);
    ASSERT_FALSE(GVL_Troubleshooting.O_MotionM2.Step8_OutputInterlockOk,
                 'M2 F4 tempos : demande retenue -> Step8 doit etre FALSE');
END_TEST

TEST 'TC-P14-TSV-15 Gate Enable/AU perdue (DISABLED) -> Step8 PAS vert'
    (* Le terme DISABLED est le SEUL qui bascule Step8 dans une situation SEMI-NOMINALE (tout est
       pret, seule la gate Enable/PowerContactorEngaged manque). Son oubli etait indetectable dans
       la v1 du garde-fou (REX revue independante T371). *)
    FB.WinchM1.State.FinalInterlockError  := FALSE;
    FB.WinchM1.State.FinalInterlockReason := E_WinchFinalInterlockReason.NONE;
    FB.WinchM1.State.FinalInterlockState  := E_WinchFinalInterlockState.DISABLED;  // :169
    FB.WinchM1.State.FinalMotorRequest    := FALSE;
    FB.WinchM1.State.BrakeCmd             := FALSE;
    FB(Enable := TRUE);
    ASSERT_FALSE(GVL_Troubleshooting.N_MotionM1.Step8_OutputInterlockOk,
                 'Gate Enable/AU perdue : etage de sortie neutralise -> Step8 doit etre FALSE');
END_TEST

TEST 'TC-P14-TSV-16 Cause MEMORISEE apres acquittement -> Step8 reste VERT (pas de faux rouge permanent)'
    (* Garde-fou de la decision A2 : `Reason` est MEMORISE et n'est pas remis a NONE quand le latch
       §3bis est acquitte (FB_WinchOutputInterlock.st:510-514). Le diagnostic doit rester VERT :
       l'injecter dans la decision produirait un faux ROUGE PERMANENT. Verifie que G522 l'interdit. *)
    FB.WinchM1.State.FinalInterlockError  := FALSE;
    FB.WinchM1.State.FinalInterlockState  := E_WinchFinalInterlockState.READY;                // latch acquitte
    FB.WinchM1.State.FinalInterlockReason := E_WinchFinalInterlockReason.SENSE_DROP_TIMEOUT;  // memoire qui reste
    FB.WinchM1.State.FinalMotorRequest    := TRUE;
    FB.WinchM1.State.RelayFwd             := TRUE;
    FB.WinchM1.State.RelayRev             := FALSE;
    FB.WinchM1.State.BrakeCmd             := TRUE;    // mouvement autorise de nouveau
    FB(Enable := TRUE);
    ASSERT_TRUE(GVL_Troubleshooting.N_MotionM1.Step8_OutputInterlockOk,
                'Cause memorisee mais barriere de nouveau autorisante -> Step8 = TRUE');
    ASSERT_EQ(GVL_Troubleshooting.N_MotionM1.Step8_InterlockReason, E_WinchFinalInterlockReason.SENSE_DROP_TIMEOUT,
              'la cause memorisee reste LISIBLE (champ de lecture) sans etre DECISIONNELLE');
END_TEST

TEST 'TC-P14-TSV-17 Vert nominal M2 et M3 -> Step8 VERT (pas de faux rouge sur les autres axes)'
    (* Couverture manquante relevee par la revue : aucun cas vert n'existait pour M2 et M3. *)
    FB.WinchM2.State.FinalInterlockError  := FALSE;
    FB.WinchM2.State.FinalInterlockReason := E_WinchFinalInterlockReason.NONE;
    FB.WinchM2.State.FinalInterlockState  := E_WinchFinalInterlockState.READY;
    FB.WinchM2.State.FinalMotorRequest    := TRUE;
    FB.WinchM2.State.RelayFwd             := TRUE;
    FB.WinchM2.State.RelayRev             := FALSE;
    FB.WinchM2.State.BrakeCmd             := TRUE;
    FB(Enable := TRUE);
    ASSERT_TRUE(GVL_Troubleshooting.O_MotionM2.Step8_OutputInterlockOk,
                'M2 nominal en mouvement -> Step8 = TRUE');

    FB.Translation.State.FinalInterlockError  := FALSE;
    FB.Translation.State.FinalInterlockState  := E_State.READY;
    FB.Translation.State.FinalInterlockReason := E_TranslationFinalInterlockReason.NONE;
    FB(Enable := TRUE);
    ASSERT_TRUE(GVL_Troubleshooting.P_MotionM3.Step8_OutputInterlockOk,
                'M3 nominal (pas de defaut) -> Step8 = TRUE');
    ASSERT_EQ(GVL_Troubleshooting.P_MotionM3.Step8_InterlockState, E_WinchFinalInterlockState.READY,
              'M3 : E_State.READY projete sur le vocabulaire commun (READY)');
END_TEST
